Fanuc KAREL source: kb00154.KL

-- PROVISIONAL review KL for V940-1; original PC SHA256 524dfa2c07804776c6e1877156dc857779b757a37636c8281a240c5e0eaa57c3
-- Incomplete behavior may be omitted. Consult companion uncertainty JSON. Do not deploy.
PROGRAM KB00154
%NOLOCKGROUP
BEGIN
  -- V9_ZERO_TABLE_METADATA_HINT layout=0002_ascii; no indexed target words; source/name/runtime held
  -- UNRESOLVED_PC offsets 5-14; opcodes 3F,75
  -- UNRESOLVED_PC offsets 19-28; opcodes 3F,75
  -- UNRESOLVED_PC offsets 33-40; opcodes 9D,23
  -- UNRESOLVED_PC offsets 45-73; opcodes 27,22,2A,22,2A,22,27,9D,31
  -- UNRESOLVED_PC offsets 78-82; opcodes 7F
END KB00154
